TYPE ST_LightCmd :
STRUCT
    eAction     : E_LightAction;
    nBrightness : UINT;
END_STRUCT
END_TYPE

(* stored: Version 1.1.0.1, ProductVersion 3.1.4026.20
   DUT ST_LightCmd: Id {D7C9A3E1-6F42-4A8D-9B31-2C5E7F901002} *)
